FUNCTION_BLOCK PositionManager (* Basic Function Block Type *)
  (* Standard: 61499-2 *)
  (* Version 0.0, 10/5/2026, Schneider Electric, Template *)
  PACKAGE SE.Nereda;
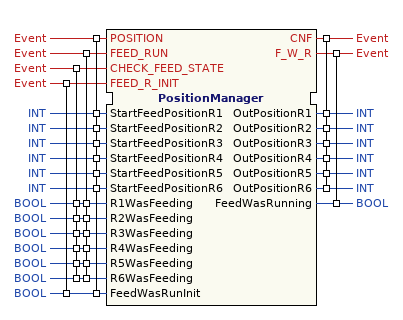
  EVENT_INPUT
    POSITION WITH StartFeedPositionR1, StartFeedPositionR2, StartFeedPositionR3, StartFeedPositionR4, StartFeedPositionR5, StartFeedPositionR6, FeedWasRunInit; (* Normal Execution Request *)
    FEED_RUN WITH R1WasFeeding, R2WasFeeding, R3WasFeeding, R4WasFeeding, R5WasFeeding, R6WasFeeding;
    CHECK_FEED_STATE WITH R1WasFeeding, R2WasFeeding, R3WasFeeding, R4WasFeeding, R5WasFeeding, R6WasFeeding;
    FEED_R_INIT WITH FeedWasRunInit;
  END_EVENT
  EVENT_OUTPUT
    CNF WITH OutPositionR1, OutPositionR2, OutPositionR3, OutPositionR4, OutPositionR5, OutPositionR6; (* Execution Confirmation *)
    F_W_R WITH FeedWasRunning;
  END_EVENT
  VAR_INPUT
    StartFeedPositionR1 : INT; (* Input event qualifier *)
    StartFeedPositionR2 : INT;
    StartFeedPositionR3 : INT;
    StartFeedPositionR4 : INT;
    StartFeedPositionR5 : INT;
    StartFeedPositionR6 : INT;
    R1WasFeeding : BOOL;
    R2WasFeeding : BOOL;
    R3WasFeeding : BOOL;
    R4WasFeeding : BOOL;
    R5WasFeeding : BOOL;
    R6WasFeeding : BOOL;
    FeedWasRunInit : BOOL;
  END_VAR
  VAR_OUTPUT
    OutPositionR1 : INT;
    OutPositionR2 : INT;
    OutPositionR3 : INT;
    OutPositionR4 : INT;
    OutPositionR5 : INT;
    OutPositionR6 : INT;
    FeedWasRunning : BOOL;
  END_VAR
  VAR
    InStartFeedPositionR1 : INT;
    InStartFeedPositionR2 : INT;
    InStartFeedPositionR3 : INT;
    InStartFeedPositionR4 : INT;
    InStartFeedPositionR5 : INT;
    InStartFeedPositionR6 : INT;
  END_VAR
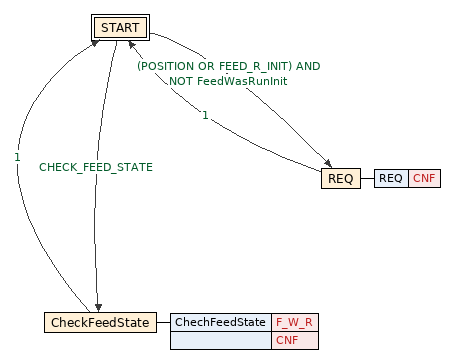
  EC_STATES
    START; (* Initial State *)
    REQ : REQ -> CNF; (* Normal execution *)
    CheckFeedState : ChechFeedState -> F_W_R, -> CNF;
  END_STATES
  EC_TRANSITIONS
    START TO CheckFeedState := CHECK_FEED_STATE;
    REQ TO START := 1;
    CheckFeedState TO START := 1;
    START TO REQ := (POSITION OR FEED_R_INIT) AND NOT FeedWasRunInit;
  END_TRANSITIONS
  ALGORITHM REQ IN ST: (* Normally executed algorithm *)
;
OutPositionR1 := StartFeedPositionR1;
OutPositionR2 := StartFeedPositionR2;
OutPositionR3 := StartFeedPositionR3;
OutPositionR4 := StartFeedPositionR4;
OutPositionR5 := StartFeedPositionR5;
OutPositionR6 := StartFeedPositionR6;
  END_ALGORITHM
  ALGORITHM ChechFeedState IN ST:
;
FeedWasRunning := R1WasFeeding OR R2WasFeeding OR R3WasFeeding OR R4WasFeeding OR R5WasFeeding OR R6WasFeeding;

IF NOT FeedWasRunning THEN
	OutPositionR1 := StartFeedPositionR1;
	OutPositionR2 := StartFeedPositionR2;
	OutPositionR3 := StartFeedPositionR3;
	OutPositionR4 := StartFeedPositionR4;
	OutPositionR5 := StartFeedPositionR5;
	OutPositionR6 := StartFeedPositionR6;
ELSE
	IF R1WasFeeding THEN
		OutPositionR1 := 1;
		OutPositionR2 := 2;
		OutPositionR3 := 0;
		OutPositionR4 := 0;
		OutPositionR5 := 0;
		OutPositionR6 := 0;
	ELSIF R2WasFeeding THEN
		OutPositionR1 := 2;
		OutPositionR2 := 1;
		OutPositionR3 := 0;
		OutPositionR4 := 0;
		OutPositionR5 := 0;
		OutPositionR6 := 0;
	END_IF;
END_IF;
  END_ALGORITHM
END_FUNCTION_BLOCK
